// TIA Portal V21 export
TagTable "T_V1"
  X_V1 :   (PLC tag HMI_IF.SwOn, HMI_Connection_1, 100 ms)
